(* PLC project zarechnaya.project, CODESYS CODESYS V3.5 SP17 Patch 3 *)
(* stored: creationDateTime 2026-10-20T05:42:22.2802919, modificationDateTime 1601-01-01T03:00:00 *)

(* FB_RatioCfc — соотношение реагента к расходу (CFC, две страницы, порядок не по схеме). Поведение (модель scenarios/reference/model_FB_RatioCfc.py), шаги executionOrderId: 1. rPrev := m — выход MUL читается раньше его шага: значение прошлого вызова (начально 0); 2. m := rFlow · rK; 3. rNow := m; 4. s := m + rBias; 5. rSum := s. Страница 1 — входы и MUL, страница 2 — сумматор и выходы. REAL (float32). *)
FUNCTION_BLOCK FB_RatioCfc
  VAR_INPUT
    rFlow : REAL;
    rK : REAL;
    rBias : REAL;
  END_VAR
  VAR_OUTPUT
    rPrev : REAL;
    rNow : REAL;
    rSum : REAL;
  END_VAR
  VAR  (* added by the conversion: wires and edge detectors of the diagram *)
    _MUL5_OUT : ANY;
  END_VAR

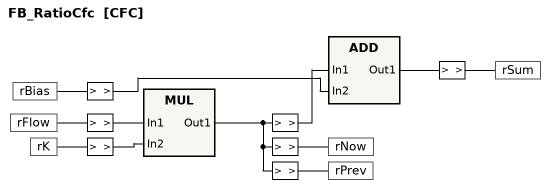
(* CFC diagram, written out as Structured Text *)
rPrev := _MUL5_OUT;
_MUL5_OUT := rFlow * rK;
rNow := _MUL5_OUT;
rSum := _MUL5_OUT + rBias;
END_FUNCTION_BLOCK
